FUNCTION_BLOCK RejectWorkpiece (* Composite Function Block Type *)
  (* Standard: 61499-2 *)
  (* Version 0.0, 7/2/2026, template *)
  PACKAGE Main;
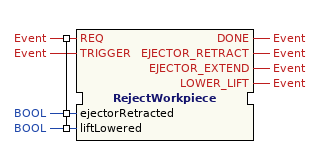
  EVENT_INPUT
    REQ WITH ejectorRetracted, liftLowered; (* Normal Execution Request *)
    TRIGGER;
  END_EVENT
  EVENT_OUTPUT
    DONE; (* Initialization Confirm *)
    EJECTOR_RETRACT; (* Execution Confirmation *)
    EJECTOR_EXTEND;
    LOWER_LIFT;
  END_EVENT
  VAR_INPUT
    ejectorRetracted : BOOL; (* Input event qualifier *)
    liftLowered : BOOL;
  END_VAR
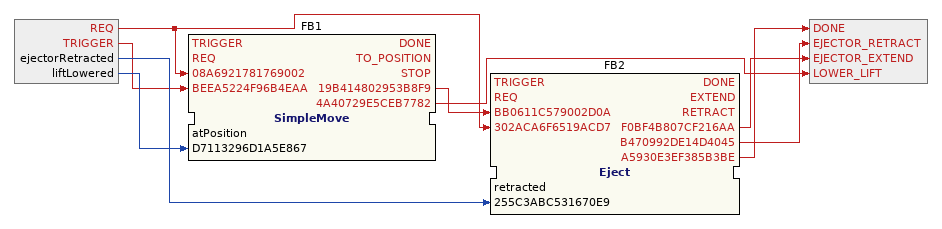
  FBS
    FB1 : SimpleMove;
    FB2 : Eject;
  END_FBS
  EVENT_CONNECTIONS
    FB2.F0BF4B807CF216AA TO EJECTOR_EXTEND;
    FB2.B470992DE14D4045 TO EJECTOR_RETRACT;
    FB2.A5930E3EF385B3BE TO DONE;
    FB1.19B414802953B8F9 TO FB2.BB0611C579002D0A;
    FB1.4A40729E5CEB7782 TO LOWER_LIFT;
    REQ TO FB2.302ACA6F6519ACD7;
    REQ TO FB1.08A6921781769002;
    TRIGGER TO FB1.BEEA5224F96B4EAA;
  END_CONNECTIONS
  DATA_CONNECTIONS
    liftLowered TO FB1.D7113296D1A5E867;
    ejectorRetracted TO FB2.255C3ABC531670E9;
  END_CONNECTIONS
END_FUNCTION_BLOCK
